Fanuc KAREL source: KD00056.KL

PROGRAM KD00056
%NOLOCKGROUP
%DEFGROUP = 1
VAR
  I: INTEGER
  J: INTEGER
  B: BOOLEAN
  R: REAL
  S: STRING[80]
  P: POSITION
BEGIN
  MOVE TO P,
  WHEN AT NODE[1] DO DOUT[1] = TRUE
  ENDMOVE
END KD00056
